// Core §10.5.1 reusable topology mechanism: bounded registration, validation,
// live value/health refresh and exact-tag diagnostic correlation.
FUNCTION_BLOCK FB_IoTopologyPublisher_Tests EXTENDS TcUnit.FB_TestSuite
VAR
    _publisher, _publisherDuplicate : FB_IoTopologyPublisher;
    _data, _dataDuplicate : ST_FieldbusTopology;
    _d : ST_Diagnostic;
    _wired, _duplicateWired : BOOL;
    // Unit rows: one table of their own, because the refused definition marks
    // its table invalid. The other two rows read only their own slots.
    _unitPublisher : FB_IoTopologyPublisher;
    _unitData : ST_FieldbusTopology;
    _unitsWired : BOOL;
END_VAR

Publishes_value_health_and_diagnostic();
Rejects_duplicate_channel_identity();
UnitCode_derives_the_unit_text();
No_code_keeps_the_catalog_text();
A_code_and_a_text_together_are_refused();

METHOD Publishes_value_health_and_diagnostic
TEST('Publishes_value_health_and_diagnostic');
IF NOT _wired THEN
    _publisher.Setup(DataRef := _data, ResetData := TRUE);
    _publisher.M_DefineNode(Index := 1, Name := 'Master',
        DescriptionKey := 'project.hardware.master', TypeId := 'Test',
        Address := 'Master', ParentIndex := 0);
    _publisher.M_DefineNode(Index := 2, Name := 'DI',
        DescriptionKey := 'project.hardware.di', TypeId := 'Test DI',
        Address := 'Terminal 1', ParentIndex := 1);
    _publisher.M_DefineDigitalChannel(NodeIndex := 2, ChannelIndex := 1,
        Tag := '_101B202A', DescriptionKey := 'project.io.101B202A',
        Address := 'EL1809 Ch5', Path := 'Unit.IO._101B202A',
        ModulePath := 'Unit.PressRam', Dir := E_ChannelDir.INPUT);
    _wired := TRUE;
END_IF
AssertTrue(Condition := _publisher.M_Validate(), Message := 'valid catalog accepted');
_publisher.M_SetAllHealth(Healthy := TRUE);
AssertTrue(Condition := _publisher.M_SetDigitalValue(
    NodeIndex := 2, ChannelIndex := 1, Value := TRUE), Message := 'known channel updated');
_d.ReasonCode := PL_ModuleReasons.CYL_NOT_EXTENDED;
_d.Description := 'project.error.pressDownSensorTimeout';
_d.IoTag := '_101B202A';
_publisher.M_BeginDiagnosticRefresh();
_publisher.M_ApplyDiagnostic(Diagnostic := _d);
AssertTrue(Condition := _data.Nodes[2].Channels[1].BoolValue,
    Message := 'live value is published');
AssertTrue(Condition := _data.Nodes[2].Channels[1].Quality,
    Message := 'aggregate health reaches the channel');
AssertTrue(Condition := _data.Nodes[2].Channels[1].FaultActive,
    Message := 'exact diagnostic tag highlights the channel');
AssertEquals_STRING(Expected := 'project.error.pressDownSensorTimeout',
    Actual := _data.Nodes[2].Channels[1].Diagnostic,
    Message := 'channel carries the diagnostic localization key');
TEST_FINISHED();
END_METHOD

METHOD Rejects_duplicate_channel_identity
TEST('Rejects_duplicate_channel_identity');
IF NOT _duplicateWired THEN
    _publisherDuplicate.Setup(DataRef := _dataDuplicate, ResetData := TRUE);
    _publisherDuplicate.M_DefineNode(Index := 1, Name := 'Master',
        DescriptionKey := 'project.hardware.master', TypeId := 'Test',
        Address := 'Master', ParentIndex := 0);
    _publisherDuplicate.M_DefineDigitalChannel(NodeIndex := 1, ChannelIndex := 1,
        Tag := '_DUPLICATE', DescriptionKey := 'project.io.first',
        Address := 'Ch1', Path := 'Unit.IO.First', ModulePath := 'Unit',
        Dir := E_ChannelDir.INPUT);
    _publisherDuplicate.M_DefineDigitalChannel(NodeIndex := 1, ChannelIndex := 2,
        Tag := '_DUPLICATE', DescriptionKey := 'project.io.second',
        Address := 'Ch2', Path := 'Unit.IO.Second', ModulePath := 'Unit',
        Dir := E_ChannelDir.INPUT);
    _duplicateWired := TRUE;
END_IF
AssertFalse(Condition := _publisherDuplicate.M_Validate(),
    Message := 'duplicate approved tag fails validation');
AssertEquals_STRING(Expected := 'std.error.fieldbusChannelIdentityDuplicate',
    Actual := _dataDuplicate.MappingDiagnostic,
    Message := 'mapping failure is explicit and localizable');
TEST_FINISHED();
END_METHOD

METHOD PRIVATE _M_WireUnits
IF _unitsWired THEN
    RETURN;
END_IF
_unitPublisher.Setup(DataRef := _unitData, ResetData := TRUE);
_unitPublisher.M_DefineNode(Index := 1, Name := 'Master',
    DescriptionKey := 'project.hardware.master', TypeId := 'Test AI',
    Address := 'Master', ParentIndex := 0);
_unitsWired := TRUE;
END_METHOD

METHOD UnitCode_derives_the_unit_text
TEST('UnitCode_derives_the_unit_text');
_M_WireUnits();
AssertTrue(Condition := _unitPublisher.M_DefineAnalogChannel(NodeIndex := 1, ChannelIndex := 1,
        Tag := '_101B301', DescriptionKey := 'project.io.101B301',
        Address := 'EL3062 Ch1', Path := 'Unit.IO._101B301',
        ModulePath := 'Unit.SupplyPressure', Dir := E_ChannelDir.INPUT,
        EngUnit := '', UnitCode := E_EngUnit.BAR),
    Message := 'a channel with a unit code is accepted');
AssertEquals_DINT(Expected := TO_DINT(E_EngUnit.BAR),
    Actual := TO_DINT(_unitData.Nodes[1].Channels[1].UnitCode),
    Message := 'the code is the published unit');
AssertEquals_STRING(Expected := 'bar', Actual := _unitData.Nodes[1].Channels[1].Unit,
    Message := 'the legacy text is derived from the code, not given twice');
TEST_FINISHED();
END_METHOD

METHOD No_code_keeps_the_catalog_text
TEST('No_code_keeps_the_catalog_text');
_M_WireUnits();
AssertTrue(Condition := _unitPublisher.M_DefineAnalogChannel(NodeIndex := 1, ChannelIndex := 2,
        Tag := '_101B302', DescriptionKey := 'project.io.101B302',
        Address := 'EL3062 Ch2', Path := 'Unit.IO._101B302',
        ModulePath := 'Unit.SupplyPressure', Dir := E_ChannelDir.INPUT,
        EngUnit := 'mA', UnitCode := E_EngUnit.NONE),
    Message := 'a unit the vocabulary lacks is given as text');
AssertEquals_DINT(Expected := TO_DINT(E_EngUnit.NONE),
    Actual := TO_DINT(_unitData.Nodes[1].Channels[2].UnitCode),
    Message := 'no code is published as NONE');
AssertEquals_STRING(Expected := 'mA', Actual := _unitData.Nodes[1].Channels[2].Unit,
    Message := 'the catalog text is kept as it is');
TEST_FINISHED();
END_METHOD

METHOD A_code_and_a_text_together_are_refused
TEST('A_code_and_a_text_together_are_refused');
_M_WireUnits();
AssertFalse(Condition := _unitPublisher.M_DefineAnalogChannel(NodeIndex := 1, ChannelIndex := 3,
        Tag := '_101B303', DescriptionKey := 'project.io.101B303',
        Address := 'EL3062 Ch3', Path := 'Unit.IO._101B303',
        ModulePath := 'Unit.SupplyPressure', Dir := E_ChannelDir.INPUT,
        EngUnit := 'psi', UnitCode := E_EngUnit.BAR),
    Message := 'two sources for one unit are a mapping defect, not resolved silently');
AssertEquals_STRING(Expected := '', Actual := _unitData.Nodes[1].Channels[3].Name,
    Message := 'the refused channel is not written');
AssertFalse(Condition := _unitData.MappingValid, Message := 'the catalog is reported invalid');
AssertEquals_STRING(Expected := 'std.error.fieldbusChannelMappingInvalid',
    Actual := _unitData.MappingDiagnostic, Message := 'with the existing mapping diagnostic');
TEST_FINISHED();
END_METHOD

END_FUNCTION_BLOCK

(* stored: Version 1.1.0.1, ProductVersion 3.1.4024.12
   POU FB_IoTopologyPublisher_Tests: Id {48966180-c90b-4d64-af4f-b1736243839f}, SpecialFunc None
   Method Publishes_value_health_and_diagnostic: Id {fc91f74a-2a63-41f2-af02-1d40e1f6b90a}
   Method Rejects_duplicate_channel_identity: Id {26c26643-487e-4ce8-8c50-8f9403b07f64}
   Method _M_WireUnits: Id {8e29905a-2ecc-4e09-ae12-776fe5c9b1c7}
   Method UnitCode_derives_the_unit_text: Id {a38d26fa-cf68-4cbd-b0f2-da3ea68580dd}
   Method No_code_keeps_the_catalog_text: Id {b27dfa43-10ac-4952-bc1c-fba5d55692e7}
   Method A_code_and_a_text_together_are_refused: Id {4dcd728f-6a9a-41ab-a138-c9bff2c6df2c} *)
